(* IEC 61131-3 sources: Lab3/Libraries/AsIOTime, 3 files *)

(* ---- AsIOTime.typ ---- *)
TYPE

END_TYPE

(* ---- AsIOTime.fun ---- *)
{REDUND_OK} {REDUND_UNREPLICABLE} FUNCTION AsIOTimeStamp : DINT (* Get current SystemTime stamp in microseconds *)
END_FUNCTION

{REDUND_CONTEXT} {REDUND_UNREPLICABLE} FUNCTION AsIOTimeCyclicStart : DINT (* Get SystemTime at start of cyclic ressource *)
END_FUNCTION

(* ---- AsIOTime.var ---- *)
VAR CONSTANT

END_VAR
